// Mitsubishi GX Works2 project: Task2_Ex_3   PLC: FX3G

PROGRAM MAIN
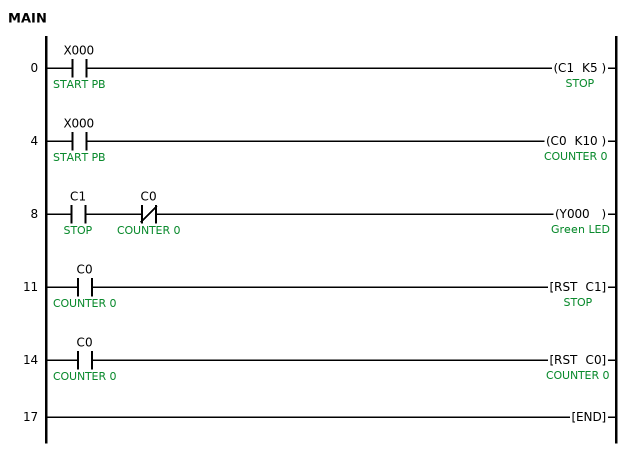
0     LD      X000  ; START PB
      OUT     C1 K5  ; STOP
4     LD      X000  ; START PB
      OUT     C0 K10  ; COUNTER 0
8     LD      C1  ; STOP
      ANI     C0  ; COUNTER 0
      OUT     Y000  ; Green LED
11    LD      C0  ; COUNTER 0
      RST     C1  ; STOP
14    LD      C0  ; COUNTER 0
      RST     C0  ; COUNTER 0
17    END
END_PROGRAM

// device comments not shown above
X001  ; RST
